// TIA Portal V20 export
// export: Created 2026-10-12T05:42:27.8855656Z, ExportSetting WithDefaults, DisplayName Totally Integrated Automation Portal, DisplayVersion V20, DisplayName TIA Portal Openness, DisplayVersion V20, DisplayName TIA Portal Teamcenter Gateway, DisplayVersion V20, DisplayName TIA Portal Version Control Interface, DisplayVersion V20, DisplayName SINAMICS Startdrive Advanced, DisplayVersion V20 SP1 Update 2, DisplayName SINAMICS Startdrive G110M, G120, G120C, G120D, G120P, G115D, DisplayVersion V20 SP1 Update 2, DisplayName SINAMICS Startdrive G130, G150, S120, S150, SINAMICS MV, G220, S200, S210, DisplayVersion V20 SP1 Update 2, DisplayName STEP 7 Professional, DisplayVersion V20, DisplayName STEP 7 Safety, DisplayVersion V20, DisplayName WinCC Basic/Comfort/Advanced, DisplayVersion V20, DisplayName WinCC Professional, DisplayVersion V20, DisplayName WinCC Unified, DisplayVersion V20
FUNCTION "FRK_SetIdentity" : Void   // FC1, SCL
{ S7_Optimized_Access := 'TRUE' }
VERSION : 0.1
// Generated registry services v0.1; compact rows contain no operator strings.
// stored: AutoNumber true, IsIECCheckEnabled false, SetENOAutomatically false, UDAEnableTagReadback false
   VAR_INPUT
      InstancePath : WString;
      ModuleType : DInt;
      TypeId : DInt;
      Capabilities : DWord;
      ParentIndex : DInt;
      TypeKey : String;
   END_VAR
   VAR_IN_OUT
      Core : "FRK_Core";
      Status : "ST_ModuleStatus";
   END_VAR
   VAR_TEMP
      Identity : String[254];
      QuotePos : Int;
      RowIndex : DInt;
   END_VAR
BEGIN

   #Core.Named := TRUE;
   #Core.RegIndex := 0;
   IF "FRK_Registry".Fault OR "FRK_Registry".Count < 0 OR "FRK_Registry".Count > 4
       OR #ParentIndex < 0 OR #ParentIndex > "FRK_Registry".Count OR #ParentIndex > 4 THEN
       "FRK_Registry".Fault := TRUE;
       RETURN;
   END_IF;
   IF #ParentIndex > 0 THEN
       IF NOT "FRK_Registry".Rows[#ParentIndex].Valid THEN
           "FRK_Registry".Fault := TRUE;
           RETURN;
       END_IF;
   END_IF;
   IF LEN(#InstancePath) > 254 THEN
       "FRK_Registry".Fault := TRUE;
       RETURN;
   END_IF;
   #Identity := WSTRING_TO_STRING(#InstancePath);
   #QuotePos := FIND(IN1 := #Identity, IN2 := '"');
   WHILE #QuotePos > 0 DO
       #Identity := DELETE(IN := #Identity, L := 1, P := #QuotePos);
       #QuotePos := FIND(IN1 := #Identity, IN2 := '"');
   END_WHILE;
   IF LEN(#Identity) > 80 OR LEN(#Identity) = 0 OR "FRK_Registry".Count >= 4 THEN
       "FRK_Registry".Fault := TRUE;
       RETURN;
   END_IF;
   "FRK_Registry".Count := "FRK_Registry".Count + 1;
   #RowIndex := "FRK_Registry".Count;
   #Core.RegIndex := #RowIndex;
   #Core.ParentIndex := #ParentIndex;
   #Core.ModuleType := #ModuleType;
   #Status.Name := #Identity;
   #Status.TypeKey := #TypeKey;
   #Status.ModuleType := #ModuleType;
   #Status.TileEnable := TRUE;
   "FRK_Registry".Rows[#RowIndex].Valid := TRUE;
   "FRK_Registry".Rows[#RowIndex].Parent := #ParentIndex;
   "FRK_Registry".Rows[#RowIndex].ModuleType := #ModuleType;
   "FRK_Registry".Rows[#RowIndex].TypeId := #TypeId;
   "FRK_Registry".Rows[#RowIndex].Capabilities := #Capabilities;
END_FUNCTION
